// Nature d'un signal de l'image E/S (docs/04 § 5)
{attribute 'qualified_only'}
{attribute 'strict'}
TYPE E_SignalKind :
(
    None := 0,
    DI := 1,
    DO := 2,
    AI := 3,
    AO := 4
) USINT;
END_TYPE

(* stored: Version 1.1.0.1, ProductVersion 3.1.4024.12
   DUT E_SignalKind: Id {3c8acf07-4291-5279-90dd-486610465aa6} *)
